(* CODESYS project teltonikaSMSalarmSender.export

Project tree, tasks and I/O mapping:
  libraries: Standard, 3.5.18.0 (System); WagoSysCurl, 1.1.5.0 (WAGO); WagoAppTime, 1.7.3.5 (WAGO); VisuDialogs, * (System)
  task MainTask (cyclic, interval 200 ms, priority 15) calls prg_AlarmSMS
  task VISU_TASK (cyclic, interval 100 ms, priority 15) calls VisuElems.Visu_Prg
  Teltonika/
    global variables GVL_TeltonikaCredentials
    function block FbAlarmSlot [ST]
    function block FbTeltonikaSMS [ST]: ExtractJson
    program prg_AlarmSMS [ST]
  visualisation AlarmAlarms
  visualisation AlarmerListe
  visualisation AlarmMain
*)

// Teltonika/GVL_TeltonikaCredentials
(*
	GVL_TeltonikaCredentials                                  Revised 22.08.2026
	==========================================================================
	WHAT THIS LIST IS FOR
	The single place where the Teltonika router login is maintained. Both the
	older prg_SendSMS and the newer prg_AlarmSMS read from here, so a
	changed password only has to be entered once.

	WHY THE CREDENTIALS ARE RETAIN AND THE REST IS NOT
	Teltonika_Username and Teltonika_Password are VAR_GLOBAL RETAIN, so they
	keep their value through a PLC restart and can be corrected online without
	rebuilding and downloading. That matters because a password change on the
	router would otherwise take a full engineering session to follow.
	The remaining entries are ordinary globals: they belong to the project and
	should come back from the source on every download.

	WHY THE PASSWORD IS BLANK IN THE SOURCE
	So the secret is not stored in the project file, which gets copied, backed
	up and shared. Enter it ONCE online and the retain keeps it.
	If you do decide to put it in the source anyway, remember that the dollar
	sign is the escape character in ST and must be doubled. Ordinary characters
	such as the at sign need no escaping.

	VERIFIED 22.08.2026 ON rutx09-hyc
	The whole API flow - login, modem status returning id 3-1, and send - works
	with the ADMIN user. A separate low privilege user named pfc300 was refused
	with HTTP 401 code 120: it either does not exist on that router, or its user
	group has no API access. To move to a dedicated API user later, create it on
	the correct router, put it in a group allowed to reach the messages
	endpoints, and change the two retain values online. No code change needed.

	Do not publish or share this file.
*)
{attribute 'qualified_only'}
VAR_GLOBAL
	// prg_AlarmSMS therefore overrides the host locally in its own
	// sRouterOverride, and only borrows the credentials from here.
	// Written WITHOUT the https prefix - the send block adds that itself.
	Teltonika_sRouterIP	: STRING := 'rutx09.tailescale.ts.net';

	// Default recipient and message for the older prg_SendSMS. The alarm
	// system does not use these; it keeps its own recipient list.
	Teltonika_Number	: STRING[64] := '+4791919191';
	Teltonika_sMessage	: STRING := 'Debug test SMSCodesys';
END_VAR

VAR_GLOBAL RETAIN
	// Router API user. Must have API rights - an ordinary low privilege user
	// is refused with 401 code 120 even when the password is correct.
	Teltonika_Username	: STRING[64] := 'admin';

	// Blank on purpose, see the note in the header. Enter it online once.
	Teltonika_Password	: STRING[64] := '';
END_VAR

// Teltonika/prg_AlarmSMS
(*
	prg_AlarmSMS                        Created 20.08.2026, rev 23.08.2026
	==========================================================================
	WHAT THIS PROGRAM DOES
	It turns boolean alarm conditions into text messages, and hands them one at
	a time to FbTeltonikaSMS, which talks to a Teltonika RUTX09 router
	over its REST API. The router holds the SIM card, so the PLC needs no modem.

	THE CHAIN, IN ORDER
	  aAlarm[i].xAlarmIn        a condition in the plant becomes TRUE
	  aAlarm[i]                 the slot debounces it and produces xActive plus
	                            the one shot edges xRising and xFalling
	  aAlarm[i].xSmsEnable      the operator switch: may this alarm send at all?
	  aAlarm[i].axToRecipient[] one BOOL per person, picking who gets this alarm
	  aQueueMsg / aQueueNo      a FIFO, because sending takes seconds and alarms
	                            can arrive in bursts
	  oSms                      the router client, driven one message at a time

	WHY EACH ALARM IS A FUNCTION BLOCK INSTANCE
	The CODESYS Best Practices for visualization recommend passing ONE parameter
	to a reusable visualization through VAR_IN_OUT. A slot instance is exactly
	that: a frame showing one row references prg_AlarmSMS.aAlarm[i] and
	gets every field of that alarm with it.

	WHY THE RECIPIENT SELECTION IS AN ARRAY OF BOOL
	Changed 23.08.2026 from a BYTE bit mask. A mask is compact but hostile to a
	visualization: a checkbox has to bind to a single bit, the operator sees a
	meaningless number, and an off by one in the bit index is invisible until
	the wrong person is woken up. One BOOL per recipient binds directly to a
	checkbox and reads the same way in the code.

	WHY A QUEUE AND A RATE LIMIT
	One message needs several task cycles and up to three network round trips.
	Without a queue a burst of alarms would overwrite each other. Without
	iMaxSmsPerHour a chattering signal could send hundreds of messages, which
	costs real money and buries the operator in noise.

	NOTE ON LANGUAGE
	Comments are English. Operator facing texts are deliberately Norwegian,
	because sText goes straight into an SMS that a Norwegian recipient reads.
*)
PROGRAM prg_AlarmSMS
VAR CONSTANT
	// Sizes are constants so the arrays, the loops and the visualization all
	// agree on one number. MAX_RECIPIENTS must match the array size declared
	// inside FbAlarmSlot - raise both together if more than four
	// people need alarms.
	MAX_ALARMS		: INT := 20;	// Alarm slots available for configuration
	MAX_RECIPIENTS	: INT := 4;		// Phone numbers that can receive alarms
	QUEUE_SIZE		: INT := 16;	// Messages that can wait before one is lost
	MAX_RETRY		: INT := 2;		// Extra attempts, and only for KNOWN failures.
									// See the retry policy in section 6 below.
	MSG_MAX_LEN		: INT := 140;	// Message cap. CONCAT returns STRING(255) in
									// CODESYS and the whole JSON body must fit in
									// that, so the text itself is capped here.
END_VAR

VAR
	// =================================================================
	// 1) THE ALARM TABLE
	// -----------------------------------------------------------------
	// One FbAlarmSlot per alarm. Each slot carries its own
	// configuration AND its own live state, and does its own debouncing.
	//
	// Wire your plant conditions into the slots from anywhere in the project:
	//   prg_AlarmSMS.aAlarm[1].xAlarmIn := NOT HTTP_HvaKosterStrommen.xPriceDataValid;
	//
	// A visualization row binds to one whole slot as a single reference:
	//   alarm  ->  prg_AlarmSMS.aAlarm[1]
	//
	// iDelaySec is in SECONDS: 30 is thirty seconds, 120 is two minutes,
	// 300 is five minutes. The slot renders it back as readable text.
	//
	// The recipient selection is NOT set here. Every slot falls back to the
	// default declared in the function block, which is recipient 1 only.
	// Change it per alarm from the visualization, or add axToRecipient to the
	// lines below if a different default suits the plant better.
	//
	// Only slots 1 to 3 are enabled. The rest are written but switched off,
	// because an alarm whose xAlarmIn is not wired yet should not be able to
	// send anything. Enable each one as you connect its signal.
	// =================================================================
	aAlarm : ARRAY[1..MAX_ALARMS] OF FbAlarmSlot := [
		// --- Energi og pris ---
		(xSmsEnable := TRUE,  iDelaySec := 300,
		 sText := 'Stroempriser ikke oppdatert fra hvakosterstrommen.no'),
		(xSmsEnable := TRUE,  iDelaySec := 120,
		 sText := 'Solcelleanlegg: ingen Modbus-kontakt'),
		(xSmsEnable := TRUE,  iDelaySec := 120,
		 sText := 'MQTT-forbindelse mot skyen er nede'),
		(xSmsEnable := FALSE, iDelaySec := 30,
		 sText := 'Hoey stroempris - forbruk boer reduseres'),

		// --- Energimaalere, stigere ---
		(xSmsEnable := FALSE, iDelaySec := 120,
		 sText := 'Energimaaler stiger 433.101 og 433.201 svarer ikke'),
		(xSmsEnable := FALSE, iDelaySec := 120,
		 sText := 'Energimaaler stiger 433.102 og 433.202 svarer ikke'),
		(xSmsEnable := FALSE, iDelaySec := 120,
		 sText := 'Energimaaler stiger 433.103 svarer ikke'),
		(xSmsEnable := FALSE, iDelaySec := 120,
		 sText := 'Energimaaler stiger 433.104 svarer ikke'),
		(xSmsEnable := FALSE, iDelaySec := 120,
		 sText := 'Energimaaler stiger 433.203 svarer ikke'),
		(xSmsEnable := FALSE, iDelaySec := 120,
		 sText := 'Energimaaler stiger 434.001 svarer ikke'),

		// --- Varme ---
		(xSmsEnable := FALSE, iDelaySec := 120,
		 sText := 'Elkjele: ingen kontakt med energimaaler'),
		(xSmsEnable := FALSE, iDelaySec := 120,
		 sText := 'Varmepumpe: ingen kontakt med energimaaler'),

		// --- Ventilasjon ---
		(xSmsEnable := FALSE, iDelaySec := 120,
		 sText := 'Ventilasjonsaggregat 360.003 svarer ikke'),
		(xSmsEnable := FALSE, iDelaySec := 120,
		 sText := 'Ventilasjonsaggregat 360.004 svarer ikke'),
		(xSmsEnable := FALSE, iDelaySec := 120,
		 sText := 'Ventilasjonsaggregat 360.005 svarer ikke'),

		// --- Varmtvann og feltbuss ---
		(xSmsEnable := FALSE, iDelaySec := 120,
		 sText := 'Varmtvannsbereder CH124 svarer ikke'),
		(xSmsEnable := FALSE, iDelaySec := 60,
		 sText := 'Modbus RTU-linje 1: kommunikasjonsfeil'),
		(xSmsEnable := FALSE, iDelaySec := 120,
		 sText := 'Teltonika-ruter: ingen Modbus-kontakt'),

		// --- Reserve ---
		(xSmsEnable := FALSE, iDelaySec := 30,
		 sText := 'Reserve - ledig alarmplass 19'),
		(xSmsEnable := FALSE, iDelaySec := 30,
		 sText := 'Reserve - ledig alarmplass 20')];

	// =================================================================
	// 2) RECIPIENTS
	// -----------------------------------------------------------------
	// Three parallel arrays, index 1 to 4. A recipient must be enabled here
	// AND selected in the slot before anything is sent, so one person can be
	// taken out of service without editing every alarm.
	//
	// In a visualization, bind a CHECKBOX to axRecipientEnable[n], and text
	// fields with %s to the name and the number.
	// =================================================================
	axRecipientEnable	: ARRAY[1..MAX_RECIPIENTS] OF BOOL       := [TRUE, FALSE, FALSE, FALSE];	// On or off per person
	asRecipientName		: ARRAY[1..MAX_RECIPIENTS] OF STRING(20) := ['Espen', '', '', ''];			// Display only, never sent
	asRecipientNumber	: ARRAY[1..MAX_RECIPIENTS] OF STRING(24) := ['+4791916159', '', '', ''];	// International format, this is what is dialled

	// =================================================================
	// 3) GENERAL SETTINGS
	// =================================================================
	xSmsGlobalEnable	: BOOL := TRUE;			// Master switch. FALSE stops all sending and all
												// queueing - use it during service work.
	xSendOkMessages		: BOOL := TRUE;			// Also send a message when an alarm clears, so the
												// operator knows the fault went away.
	sSiteName			: STRING(20) := 'PFC300';	// Prefix in every message. Essential when one
												// phone receives alarms from several plants.
	iMaxSmsPerHour		: INT := 15;			// Hard ceiling per rolling hour, against runaway cost
	tPauseBetweenSms	: TIME := T#10S;		// Gap between messages. Gives the router time to hand
												// the previous one over, and guarantees a clean edge.
	tRetryDelay			: TIME := T#60S;		// Wait before repeating a message that failed for a
												// known reason, so a brief outage can recover.

	// Leave EMPTY to fall back
	// to GVL_TeltonikaCredentials.Teltonika_sRouterIP.
	sRouterOverride		: STRING(80) := '';

	// Modem id inside the router. Leave EMPTY for auto-detection, which is
	// normal and survives the id changing after a router restart.
	sModemIdForced		: STRING(16) := '';

	// =================================================================
	// STATUS AND DIAGNOSTICS
	// -----------------------------------------------------------------
	// Read only. These exist to be bound to a visualization, and to make a
	// failure explain itself without a debugger attached.
	// =================================================================
	sRouterInUse			: STRING(80);	// Host actually used, after the override is resolved
	xCredentialsMissing		: BOOL;			// TRUE when user name or password is blank. Blocks
											// sending so the queue is not burned on doomed logins.
	iQueueCount				: INT;			// Messages waiting right now
	xRateLimited			: BOOL;			// TRUE when the hourly ceiling holds messages back
	iSentThisHour			: INT;			// Counter behind the ceiling, reset once an hour
	iEnabledCount			: INT;			// How many of the twenty alarms are switched on. Handy
											// as a single number on an overview screen.
	iActiveCount			: INT;			// How many alarms are standing right now
	udiSentOk				: UDINT;		// Messages the router confirmed, since PLC start
	udiSendFailed			: UDINT;		// Messages given up on after all allowed retries
	udiUncertain			: UDINT;		// Messages whose fate is unknown - the request went out
											// but no answer came back. Never retried, to avoid
											// sending the same SMS twice.
	udiDropped				: UDINT;		// Messages never queued because the FIFO was full
	sLastMessage			: STRING(140);	// Exact text last handed to the router
	sLastError				: STRING(200);	// Why the last attempt failed
	sSmsStatus				: STRING(200);	// Live progress text from the send FB
	sCurlError				: STRING(200);	// Raw libcurl error. The one to read when diHttpCode
											// stays 0, because then there is no HTTP answer.
	diHttpCode				: DINT;			// HTTP status of the last request. 0 means the request
											// never produced an HTTP answer at all.
	uiSendStep				: UINT;			// Live step inside the send FB: 10 and 11 login,
											// 20 and 21 modem lookup, 30 and 31 the send itself.

	// =================================================================
	// MANUAL TEST
	// -----------------------------------------------------------------
	// One button, two destinations. Leave sTestNumber EMPTY and the test goes
	// to every enabled recipient, which proves the real alarm path end to end.
	// Type a number into sTestNumber and it goes only there, which is how you
	// check a new phone before adding it to the recipient list.
	// xManualSend is self resetting, so a visualization button only has to
	// toggle it and the program clears it again on the next cycle.
	// =================================================================
	xManualSend			: BOOL;								// Set TRUE to queue one test message
	sTestNumber			: STRING(24) := '';					// Optional. Empty means all enabled recipients.
	sManualText			: STRING(100) := 'Testmelding fra PFC300';	// Body of the test message
	iTestQueued			: INT;								// How many messages the last test queued,
															// so the operator sees it did something

	// =================================================================
	// INTERNALS - not intended for the visualization
	// =================================================================
	aQueueMsg			: ARRAY[1..QUEUE_SIZE] OF STRING(140);	// FIFO slot: the message text
	aQueueNo			: ARRAY[1..QUEUE_SIZE] OF STRING(24);	// FIFO slot: the recipient number.
																// Kept beside the text so one alarm
																// to three people becomes three
																// independent queue entries.
	iQHead				: INT;					// Last slot read from, wraps at QUEUE_SIZE
	iQTail				: INT;					// Last slot written to, wraps at QUEUE_SIZE

	oSms				: FbTeltonikaSMS;	// The router client. Called every cycle so its
													// asynchronous transfer can advance.
	xSendTrigger		: BOOL;					// Rising edge starts oSms. Held TRUE for the whole
												// job and cleared afterwards, so the next message
												// gets a fresh edge.
	iSendState			: INT;					// Sender state machine, see section 6
	iRetry				: INT;					// Attempts already used on the current message
	sCurMsg				: STRING(140);			// The message being sent right now
	sCurNo				: STRING(24);			// The recipient it is going to

	TON_Pause			: TON;					// Enforces tPauseBetweenSms between messages
	TON_Retry			: TON;					// Enforces tRetryDelay before a repeat attempt
	TON_HourWindow		: TON;					// Free running one hour timer that clears
												// iSentThisHour, implementing the rate limit

	xManualPrev			: BOOL;					// Edge memory for xManualSend
	i					: INT;					// Loop counter over the alarm slots
	iRcp				: INT;					// Loop counter over the recipients. NOTE: a bare
												// r cannot be used as an identifier - CODESYS
												// reserves R and S as the IL reset and set
												// operators, and the parser fails cryptically.
	iGuard				: INT;					// Safety counter so the sanitize loop can never
												// spin forever on malformed text
	iQuote				: INT;					// Position of the next double quote to remove
	xQueueIt			: BOOL;					// Set when the slot being scanned needs sending
	sMsg				: STRING(140);			// Message being assembled
	sStamp				: STRING(30);			// Time stamp for the message, format dd.mm hh:mm
	sRaw				: STRING(40);			// Raw DT_TO_STRING output the stamp is cut from
END_VAR

// =====================================================================
// 1) Resolve which router host to talk to.
//    The local override wins, or if it is emty use so GVL_TeltonikaCredentials.Teltonika_sRouterIP
// =====================================================================
IF LEN(sRouterOverride) > 0 THEN
	sRouterInUse := sRouterOverride;
ELSE
	sRouterInUse := GVL_TeltonikaCredentials.Teltonika_sRouterIP;
END_IF

// Without credentials every login is doomed, and each doomed attempt costs a
// network round trip and fills the diagnostics with noise. Detect it once here
// and let section 6 hold the queue instead.
xCredentialsMissing := (LEN(GVL_TeltonikaCredentials.Teltonika_Username) = 0)
					OR (LEN(GVL_TeltonikaCredentials.Teltonika_Password) = 0);

// =====================================================================
// 2) Rolling one hour window behind the rate limit.
//    A free running timer is enough: it does not matter exactly where the
//    hour boundary falls, only that the counter cannot grow forever.
// =====================================================================
TON_HourWindow(IN := TRUE, PT := T#1H);
IF TON_HourWindow.Q THEN
	TON_HourWindow(IN := FALSE);	// Restart the window
	iSentThisHour := 0;
END_IF

// =====================================================================
// 3) Build the time stamp that goes into every message.
//    DT_TO_STRING has a fixed layout, so the parts can be cut out by
//    position instead of parsed:
//        DT#2026-08-20-14:20:28
//            ^4      ^9 ^12 ^15
// =====================================================================
sRaw   := DT_TO_STRING(WagoAppTime.FuGetLocalDateAndTime());
sStamp := CONCAT(MID(sRaw, 2, 12), '.');		// Two digits of day
sStamp := CONCAT(sStamp, MID(sRaw, 2, 9));		// Two digits of month
sStamp := CONCAT(sStamp, ' ');
sStamp := CONCAT(sStamp, MID(sRaw, 5, 15));		// Five characters, hh:mm

// =====================================================================
// 4) Scan every alarm slot and queue messages for the transitions.
//    Calling the slot updates its debounce timer and its edge outputs, so
//    all the per alarm timing logic lives in the slot rather than here.
//    Only transitions produce messages: a standing alarm stays silent.
// =====================================================================
iEnabledCount := 0;
iActiveCount  := 0;

FOR i := 1 TO MAX_ALARMS DO

	aAlarm[i]();			// Debounce and edge detection happen inside the slot
	xQueueIt := FALSE;

	// Two counters for the overview screen, so the operator can see at a
	// glance how much of the system is armed and how much is in alarm.
	IF aAlarm[i].xSmsEnable THEN
		iEnabledCount := iEnabledCount + 1;
	END_IF
	IF aAlarm[i].xActive THEN
		iActiveCount := iActiveCount + 1;
	END_IF

	IF xSmsGlobalEnable AND aAlarm[i].xSmsEnable THEN
		IF aAlarm[i].xRising THEN
			// The alarm has just appeared.
			sMsg     := CONCAT(sSiteName, ' ');
			sMsg     := CONCAT(sMsg, sStamp);
			sMsg     := CONCAT(sMsg, ' ALARM: ');
			sMsg     := CONCAT(sMsg, aAlarm[i].sText);
			xQueueIt := TRUE;
		ELSIF aAlarm[i].xFalling AND xSendOkMessages THEN
			// The alarm has cleared. Optional, because on a noisy signal this
			// doubles the number of messages.
			sMsg     := CONCAT(sSiteName, ' ');
			sMsg     := CONCAT(sMsg, sStamp);
			sMsg     := CONCAT(sMsg, ' OK: ');
			sMsg     := CONCAT(sMsg, aAlarm[i].sText);
			xQueueIt := TRUE;
		END_IF
	END_IF

	IF xQueueIt THEN
		// The message is embedded in a JSON body, where a double quote would
		// end the string early and corrupt the request. Replace any with
		// spaces. The guard counter bounds the loop so malformed text can
		// never stall the task.
		iGuard := 0;
		iQuote := FIND(sMsg, '"');
		WHILE (iQuote > 0) AND (iGuard < 20) DO
			sMsg   := REPLACE(sMsg, ' ', 1, iQuote);
			iQuote := FIND(sMsg, '"');
			iGuard := iGuard + 1;
		END_WHILE

		IF LEN(sMsg) > MSG_MAX_LEN THEN
			sMsg := LEFT(sMsg, MSG_MAX_LEN);
		END_IF

		// One queue entry per selected recipient. Two conditions have to agree:
		// the person must be in service at all (axRecipientEnable) AND this
		// particular alarm must be addressed to them (axToRecipient). Queueing
		// per recipient rather than per alarm keeps the sender simple: it never
		// has to know that one alarm can have several destinations.
		FOR iRcp := 1 TO MAX_RECIPIENTS DO
			IF axRecipientEnable[iRcp]
				AND aAlarm[i].axToRecipient[iRcp]
				AND (LEN(asRecipientNumber[iRcp]) > 0) THEN

				IF iQueueCount < QUEUE_SIZE THEN
					iQTail            := (iQTail MOD QUEUE_SIZE) + 1;	// Ring buffer wrap
					aQueueMsg[iQTail] := sMsg;
					aQueueNo[iQTail]  := asRecipientNumber[iRcp];
					iQueueCount       := iQueueCount + 1;
				ELSE
					// Queue full. Counting the loss is better than blocking the
					// task or discarding it unnoticed.
					udiDropped := udiDropped + 1;
				END_IF
			END_IF
		END_FOR
	END_IF
END_FOR

// =====================================================================
// 5) Manual test message.
//    Two destinations from one button:
//      sTestNumber empty     -> every enabled recipient, which proves the
//                               real alarm path exactly as an alarm would use it
//      sTestNumber filled in -> only that number, for checking a new phone
//                               before it is added to the recipient list
//    iTestQueued reports back how many messages were actually queued, so a
//    press that produced nothing is visible rather than silent.
// =====================================================================
IF xManualSend AND NOT xManualPrev THEN
	sMsg := CONCAT(sSiteName, ' ');
	sMsg := CONCAT(sMsg, sStamp);
	sMsg := CONCAT(sMsg, ' TEST: ');
	sMsg := CONCAT(sMsg, sManualText);

	// Same sanitizing as a real alarm, because the operator types this text
	// and a double quote would corrupt the JSON body just the same.
	iGuard := 0;
	iQuote := FIND(sMsg, '"');
	WHILE (iQuote > 0) AND (iGuard < 20) DO
		sMsg   := REPLACE(sMsg, ' ', 1, iQuote);
		iQuote := FIND(sMsg, '"');
		iGuard := iGuard + 1;
	END_WHILE

	IF LEN(sMsg) > MSG_MAX_LEN THEN
		sMsg := LEFT(sMsg, MSG_MAX_LEN);
	END_IF

	iTestQueued := 0;

	IF LEN(sTestNumber) > 0 THEN
		// A number was typed in, so send only there.
		IF iQueueCount < QUEUE_SIZE THEN
			iQTail            := (iQTail MOD QUEUE_SIZE) + 1;
			aQueueMsg[iQTail] := sMsg;
			aQueueNo[iQTail]  := sTestNumber;
			iQueueCount       := iQueueCount + 1;
			iTestQueued       := 1;
		ELSE
			udiDropped := udiDropped + 1;
		END_IF
	ELSE
		// No number typed, so send to everyone who is enabled - the same set
		// an alarm addressed to all four recipients would reach.
		FOR iRcp := 1 TO MAX_RECIPIENTS DO
			IF axRecipientEnable[iRcp] AND (LEN(asRecipientNumber[iRcp]) > 0) THEN
				IF iQueueCount < QUEUE_SIZE THEN
					iQTail            := (iQTail MOD QUEUE_SIZE) + 1;
					aQueueMsg[iQTail] := sMsg;
					aQueueNo[iQTail]  := asRecipientNumber[iRcp];
					iQueueCount       := iQueueCount + 1;
					iTestQueued       := iTestQueued + 1;
				ELSE
					udiDropped := udiDropped + 1;
				END_IF
			END_IF
		END_FOR
	END_IF
END_IF
xManualPrev := xManualSend;
xManualSend := FALSE;			// Clear it again so the button is momentary

// =====================================================================
// 6) The sender.
//    Strictly one message at a time. The send FB can only handle one job, and
//    serialising here also means the router is never hit by parallel requests.
//
//    RETRY POLICY, and why it is not simply MAX_RETRY attempts:
//    Repeating a request is only safe when we KNOW nothing was sent. A login
//    failure, or a rejection carrying a real HTTP status, both mean the router
//    did nothing, so those are retried. But if the send request went out and
//    no answer came back, the router may already have queued the SMS -
//    repeating it would deliver the same message twice. The send FB flags that
//    case with xSendUncertain, and such a message is dropped and counted.
// =====================================================================
CASE iSendState OF

	// -----------------------------------------------------------------
	0:	// Idle. Take the next message out of the queue if everything allows it.
	// -----------------------------------------------------------------
		xSendTrigger := FALSE;
		xRateLimited := (iSentThisHour >= iMaxSmsPerHour) AND (iQueueCount > 0);

		IF (iQueueCount > 0)
			AND xSmsGlobalEnable
			AND NOT xRateLimited
			AND NOT xCredentialsMissing THEN

			iQHead      := (iQHead MOD QUEUE_SIZE) + 1;		// Ring buffer wrap
			sCurMsg     := aQueueMsg[iQHead];
			sCurNo      := aQueueNo[iQHead];
			iQueueCount := iQueueCount - 1;
			iRetry      := 0;
			iSendState  := 10;
		END_IF

	// -----------------------------------------------------------------
	10:	// Start one attempt. Raising xSendTrigger gives the send FB the rising
	//     edge it needs; it stays TRUE until the job finishes.
	// -----------------------------------------------------------------
		sLastMessage := sCurMsg;
		xSendTrigger := TRUE;
		iSendState   := 20;

	// -----------------------------------------------------------------
	20:	// Wait for the verdict. The send FB is asynchronous and advances one
	//     step per call, so this state is held for several cycles.
	// -----------------------------------------------------------------
		IF oSms.xDone THEN
			xSendTrigger  := FALSE;
			udiSentOk     := udiSentOk + 1;
			iSentThisHour := iSentThisHour + 1;
			iSendState    := 30;

		ELSIF oSms.xError THEN
			xSendTrigger := FALSE;
			sLastError   := oSms.sErrorText;

			IF oSms.xSendUncertain THEN
				// Unknown outcome, see the retry policy above. The hour slot is
				// counted as used as well, because the message probably did cost
				// an SMS and the rate limit should not underestimate usage.
				udiUncertain  := udiUncertain + 1;
				iSentThisHour := iSentThisHour + 1;
				iSendState    := 30;

			ELSIF iRetry < MAX_RETRY THEN
				// Known failure, nothing was sent, so trying again is safe.
				iRetry     := iRetry + 1;
				iSendState := 40;

			ELSE
				// Out of attempts. Give up on this one and move on, rather than
				// letting a single bad message block the whole queue.
				udiSendFailed := udiSendFailed + 1;
				iSendState    := 30;
			END_IF
		END_IF

	// -----------------------------------------------------------------
	30:	// Pause between messages. Two purposes: breathing room for the router,
	//     and it guarantees at least one cycle with xSendTrigger FALSE so the
	//     next message produces a genuine rising edge.
	// -----------------------------------------------------------------
		TON_Pause(IN := TRUE, PT := tPauseBetweenSms);
		IF TON_Pause.Q THEN
			TON_Pause(IN := FALSE);
			iSendState := 0;
		END_IF

	// -----------------------------------------------------------------
	40:	// Wait before repeating the same message, so a brief outage has time
	//     to clear instead of burning all attempts in a few seconds.
	// -----------------------------------------------------------------
		TON_Retry(IN := TRUE, PT := tRetryDelay);
		IF TON_Retry.Q THEN
			TON_Retry(IN := FALSE);
			iSendState := 10;
		END_IF

ELSE
	// Unknown state. Reached only after an online change moves the code under
	// a running state machine. Returning to idle is always safe.
	iSendState := 0;
END_CASE

// =====================================================================
// 7) Call the router client.
//    This MUST run every cycle, including when idle: the underlying cURL
//    transfer is asynchronous and only advances when the FB body executes.
// =====================================================================
oSms(
	sRouterIP      := sRouterInUse,
	sUsername      := GVL_TeltonikaCredentials.Teltonika_Username,
	sPassword      := GVL_TeltonikaCredentials.Teltonika_Password,
	sNumber        := sCurNo,
	sMessage       := sCurMsg,
	sModemIdForced := sModemIdForced,
	xSend          := xSendTrigger);

// Mirror the interesting outputs so a visualization can bind them here rather
// than reaching into the FB instance. Everything else is still reachable as
// oSms.<name>, for example oSms.udiLoginCnt and oSms.xTokenValid.
sSmsStatus := oSms.sStatus;
sCurlError := oSms.sCurlError;		// The one that explains a diHttpCode of 0
diHttpCode := oSms.diHttpCode;
uiSendStep := oSms.uiStepOut;		// 10 and 11 login, 20 and 21 modem, 30 and 31 send

END_PROGRAM

// Teltonika/FbTeltonikaSMS
(*
	FbTeltonikaSMS                      Created 20.08.2026, rev 22.08.2026
	==========================================================================
	WHAT THIS BLOCK DOES
	Sends ONE text message through a Teltonika RUTX router using its REST API.
	The router holds the SIM card, so the PLC needs no modem. Give it a number
	and a text, pulse xSend, and watch xDone or xError.

	Reference implementation: github.com/espenbo/wagoEdgeStart/TeltonikaRouter
	and the working /root/sendsms_busyboxV3.sh on this PLC. Both were used to
	prove the API flow before it was written in ST.

	THE API FLOW - THREE REQUESTS
	  1  POST /api/login                 user and password  ->  bearer token
	  2  GET  /api/modems/status         token              ->  modem id, 3-1 here
	  3  POST /api/messages/actions/send token, number, text, modem id
	The router answers the third with success true when it has accepted the SMS.

	*** WHY EVERY REQUEST IS SPLIT IN TWO STEPS ***
	WagoSysCurl.FbCurl is ASYNCHRONOUS. curl_easy_perform() only STARTS the
	transfer and returns immediately; the FB reports progress through xBusy,
	xDone and xError, and its body must be called every cycle for those to
	update. Reading curl_easy_getResponseCode() straight after perform therefore
	always yields 0 and an empty receive buffer - which looks exactly like a
	network failure and is extremely misleading. Each request is consequently a
	start step followed by a wait step:

	  10 login start   11 login wait
	  20 modem start   21 modem wait
	  30 send start    31 send wait
	 100 done         900 error

	Every wait step is bounded by tWaitTimeout, so a transfer that never
	completes cannot freeze the state machine.

	*** TOKEN CACHING ***
	The router reports expires 299, so a token is good for just under five
	minutes. Both the token and the detected modem id survive between messages,
	so a follow up message jumps straight to step 30: two steps and one network
	round trip instead of eight steps and three. If the router rejects a cached
	token with HTTP 401 the block logs in again once and repeats the request,
	which is safe because a 401 proves nothing was sent.

	*** DUPLICATE PROTECTION ***
	If the send request goes out and no answer comes back, the router may
	already have accepted the SMS. Repeating it would deliver the same message
	twice. That case raises xSendUncertain, and the caller must not retry while
	it is set. A clean HTTP answer reporting failure is safe to repeat.

	*** LENGTH LIMITS TO RESPECT ***
	CONCAT returns STRING(255) in CODESYS, so the assembled JSON body cannot
	exceed that. sMessage is therefore capped at 140 characters, which also
	keeps the SMS inside a single 160 character GSM message.
*)
FUNCTION_BLOCK FbTeltonikaSMS
VAR_INPUT
	// --- What to send, and where ---
	sRouterIP		: STRING(80);		// Router host name or IP. WITHOUT the https prefix,
										// the block adds that when building the URL.
	sUsername		: STRING(64);		// Router API user. Must have API rights - an ordinary
										// low privilege user is rejected with 401 code 120.
	sPassword		: STRING(64);		// Password for that user
	sNumber			: STRING(32);		// Recipient, international format, for example +47...
	sMessage		: STRING(140);		// The text itself. See the length note in the header.

	// --- Behaviour tuning ---
	sModemIdForced	: STRING(16) := '';	// Leave EMPTY for auto-detection, which is normal and
										// survives the id changing after a router restart.
										// Set it only to pin one specific modem.
	tRequestTimeout	: TIME := T#15S;	// Passed down to cURL as its own transfer timeout
	tWaitTimeout	: TIME := T#30S;	// Guard in the wait steps. Keep it LONGER than
										// tRequestTimeout, so cURL gets to fail on its own
										// terms first and can report a proper reason.
	tTokenLifetime	: TIME := T#4M;		// How long a token is reused before logging in again.
										// The router says 299 s, so stay safely below that.

	// --- Control ---
	xSend			: BOOL;				// RISING EDGE starts one send job. Level is ignored
										// while a job is already running.
END_VAR
VAR_OUTPUT
	// --- Job state ---
	xBusy			: BOOL;				// TRUE from the rising edge until done or failed
	xDone			: BOOL;				// Latched TRUE when the router confirmed the SMS.
										// Cleared when the next job starts.
	xError			: BOOL;				// Latched TRUE when the job failed. Read sErrorText.
	xSendUncertain	: BOOL;				// TRUE when the SMS may or may not have gone out.
										// The caller MUST NOT retry the message while set,
										// or the recipient can receive it twice.
	xTokenValid		: BOOL;				// TRUE while a cached token can still be reused

	// --- Human readable status ---
	sErrorText		: STRING(200);		// Why the last job failed, including HTTP code and,
										// where useful, the raw answer from the router
	sStatus			: STRING(200);		// Live progress text, useful on a visualization
	tLastSend		: DT;				// Time stamp of the last confirmed send

	// --- Counters, all since PLC start ---
	sModemID		: STRING(16);		// Modem id currently in use. Kept between messages so
										// the lookup runs once rather than every time.
	udiSentCnt		: UDINT;			// Messages the router confirmed
	udiErrorCnt		: UDINT;			// Jobs that ended in failure
	udiLoginCnt		: UDINT;			// Actual logins performed. Compare with udiSentCnt to
										// see token caching working: it should stay well below.

	// --- Raw diagnostics from the last completed request ---
	diHttpCode		: DINT;				// HTTP status. 0 is special: it means the transfer
										// never produced an HTTP answer at all, so look at
										// sCurlError instead of trying to interpret the code.
	xCurlError		: BOOL;				// libcurl reported a transport level error
	sCurlError		: STRING(200);		// libcurl error text. The real explanation whenever
										// diHttpCode is 0, for example a name resolution
										// failure or an SSL connect error.
	sCurlSource		: STRING(100);		// Where inside libcurl the error came from
	sLastResponse	: STRING(200);		// First 200 characters of the router answer, so a
										// rejection can be read without a network trace
	uiStepOut		: UINT;				// Mirror of the internal step, for commissioning
END_VAR
VAR
	fbCurl			: WagoSysCurl.FbCurl;	// The cURL handle. ASYNCHRONOUS - see header.
	uiStep			: UINT;				// State machine position, see the header for the map
	xSendPrev		: BOOL;				// Edge memory for xSend
	TON_Wait		: TON;				// Bounds each wait step, so a stalled transfer cannot
										// hold the state machine forever
	TON_TokenAge	: TON;				// Ages the cached token out after tTokenLifetime
	xRetriedLogin	: BOOL;				// Allows exactly ONE forced re-login per job after a
										// 401, so a stale token cannot cause an endless loop
	sResponse		: STRING(4095);		// Receive buffer for the HTTP body. Deliberately large:
										// the modem status answer carries many fields.
	sURL			: STRING(200);		// Assembled request URL
	sBody			: STRING(254);		// Assembled JSON request body. Sized just under the
										// 255 characters CONCAT can produce.
	sHeader			: STRING(250);		// Assembled Authorization header
	sToken			: STRING(200);		// Bearer token. Reused across messages until it ages
										// out or the router rejects it.
END_VAR

// =====================================================================
// The FB body must run EVERY cycle, idle or not. The cURL transfer is
// asynchronous and only makes progress when this executes; skipping it
// would leave xBusy, xDone and xError frozen at their old values.
// =====================================================================
fbCurl();
uiStepOut := uiStep;

// =====================================================================
// Age the cached token out.
// The timer runs only while a token is held, so it measures the age of that
// specific token. When it expires the token is discarded and the next job
// logs in again. tTokenLifetime sits below the 299 seconds the router
// reports, so we never present a token the router has already forgotten.
// =====================================================================
TON_TokenAge(IN := xTokenValid, PT := tTokenLifetime);
IF TON_TokenAge.Q THEN
	xTokenValid := FALSE;
	sToken      := '';
END_IF

// =====================================================================
// A rising edge on xSend starts one job. A job in progress is never
// interrupted, so a caller cannot corrupt a transfer by pulsing again.
//
// The entry point depends on what is still cached. With a valid token and a
// known modem id the job starts directly at the send step, which is the whole
// point of the caching: two steps instead of eight.
// =====================================================================
IF xSend AND NOT xSendPrev AND NOT xBusy THEN
	xBusy          := TRUE;
	xDone          := FALSE;
	xError         := FALSE;
	xSendUncertain := FALSE;
	xRetriedLogin  := FALSE;	// Fresh job, so the one allowed re-login is available again
	sErrorText     := '';
	diHttpCode     := 0;

	IF xTokenValid AND (LEN(sToken) > 0) THEN
		IF LEN(sModemIdForced) > 0 THEN
			sModemID := sModemIdForced;
			uiStep   := 30;		// Token cached and modem pinned by the operator
		ELSIF LEN(sModemID) > 0 THEN
			uiStep   := 30;		// Token cached and modem detected earlier
		ELSE
			uiStep   := 20;		// Token cached but the modem is still unknown
		END_IF
	ELSE
		uiStep := 10;			// No usable token, so start with a login
	END_IF
END_IF
xSendPrev := xSend;

// =====================================================================
// The state machine.
//
// libcurl option numbers used below, since the WAGO wrapper takes raw ints:
//   13 = TIMEOUT in seconds     47 = POST             64 = SSL_VERIFYPEER
//   78 = CONNECTTIMEOUT         80 = HTTPGET          81 = SSL_VERIFYHOST
//   10002 = URL   10015 = POSTFIELDS   10018 = USERAGENT   10023 = HTTPHEADER
//
// Certificate checking is switched off because the router presents a self
// signed certificate that no public CA vouches for. That is acceptable here
// because the traffic already runs inside the Tailscale tunnel, which does
// its own authentication and encryption.
// =====================================================================
CASE uiStep OF

	// -----------------------------------------------------------------
	0:	// Idle, waiting for a rising edge on xSend.
	// -----------------------------------------------------------------
		xBusy := FALSE;

	// -----------------------------------------------------------------
	10:	// LOGIN - start the request.
	//     Any previous token is dropped first, so a failure here cannot leave
	//     a half valid credential behind for the next job to trip over.
	// -----------------------------------------------------------------
		sStatus     := 'Steg 10: logger inn paa ruteren...';
		sResponse   := '';
		xTokenValid := FALSE;
		sToken      := '';

		fbCurl.curl_easy_init();
		fbCurl.curl_set_RAM(ADR(sResponse), SIZEOF(sResponse));		// Where the answer lands
		fbCurl.curl_easy_setopt_BOOL(64, FALSE);					// Do not verify the certificate
		fbCurl.curl_easy_setopt_BOOL(81, FALSE);					// Do not verify the host name
		fbCurl.curl_easy_setopt_DINT(13, TIME_TO_DINT(tRequestTimeout) / 1000);
		fbCurl.curl_easy_setopt_DINT(78, 10);						// Connect timeout, seconds
		fbCurl.curl_easy_setopt_DINT(47, 1);						// This is a POST

		sURL := CONCAT('https://', sRouterIP);
		sURL := CONCAT(sURL, '/api/login');
		fbCurl.curl_easy_setopt_STRING(10002, sURL);

		// The API only accepts JSON, so the content type has to be declared.
		fbCurl.curl_slist_append(1, 'Content-Type: application/json');
		fbCurl.curl_easy_setopt_slist(10023, 1);

		sBody := CONCAT('{"username":"', sUsername);
		sBody := CONCAT(sBody, '","password":"');
		sBody := CONCAT(sBody, sPassword);
		sBody := CONCAT(sBody, '"}');
		fbCurl.curl_easy_setopt_STRING(10015, sBody);

		fbCurl.curl_easy_perform();		// Starts the transfer and returns at once
		TON_Wait(IN := FALSE);			// Arm the guard timer for the wait step
		uiStep := 11;

	// -----------------------------------------------------------------
	11:	// LOGIN - wait for the answer, then pull the token out of it.
	// -----------------------------------------------------------------
		TON_Wait(IN := TRUE, PT := tWaitTimeout);
		IF fbCurl.xDone OR fbCurl.xError THEN
			TON_Wait(IN := FALSE);

			// Capture everything libcurl knows BEFORE cleaning the handle up,
			// otherwise the diagnostics are lost with it.
			diHttpCode    := LINT_TO_DINT(fbCurl.curl_easy_getResponseCode());
			xCurlError    := fbCurl.xError;
			sCurlError    := fbCurl.sErrorString;
			sCurlSource   := fbCurl.sErrorSource;
			sLastResponse := LEFT(sResponse, 200);

			// Free the header list and the handle. Skipping this leaks memory
			// and lets headers accumulate across requests.
			fbCurl.curl_slist_free_all(1);
			fbCurl.curl_easy_cleanup();

			sToken := ExtractJson(sSource := sResponse, sKey := '"token"');
			IF LEN(sToken) > 0 THEN
				xTokenValid := TRUE;			// Also starts the token age timer
				udiLoginCnt := udiLoginCnt + 1;
				sStatus     := 'Token mottatt';
				IF LEN(sModemIdForced) > 0 THEN
					sModemID := sModemIdForced;
					uiStep   := 30;
				ELSIF LEN(sModemID) > 0 THEN
					uiStep   := 30;
				ELSE
					uiStep   := 20;
				END_IF
			ELSE
				// No token in the answer. Report the HTTP code, and add whichever
				// detail actually explains it: the router answer when there is
				// one, the libcurl reason when the transfer never got that far.
				sErrorText := CONCAT('Innlogging feilet, HTTP ', DINT_TO_STRING(diHttpCode));
				IF diHttpCode = 0 THEN
					sErrorText := CONCAT(sErrorText, ' curl: ');
					sErrorText := CONCAT(sErrorText, LEFT(sCurlError, 110));
				ELSE
					sErrorText := CONCAT(sErrorText, ' svar: ');
					sErrorText := CONCAT(sErrorText, LEFT(sResponse, 110));
				END_IF
				uiStep := 900;
			END_IF

		ELSIF TON_Wait.Q THEN
			// The transfer never reported completion. Abort it explicitly so
			// libcurl releases the connection instead of leaving it dangling.
			TON_Wait(IN := FALSE);
			fbCurl.curl_easy_abort();
			fbCurl.curl_slist_free_all(1);
			fbCurl.curl_easy_cleanup();
			sErrorText := 'Tidsavbrudd under innlogging';
			uiStep     := 900;
		END_IF

	// -----------------------------------------------------------------
	20:	// MODEM ID - start the request.
	//     The send endpoint needs to know which modem to use, and the id is
	//     not fixed: it depends on the hardware slot and can change after a
	//     router restart. Asking is more robust than hard coding.
	// -----------------------------------------------------------------
		sStatus   := 'Steg 20: henter modem-ID...';
		sResponse := '';

		fbCurl.curl_easy_init();
		fbCurl.curl_set_RAM(ADR(sResponse), SIZEOF(sResponse));
		fbCurl.curl_easy_setopt_BOOL(64, FALSE);
		fbCurl.curl_easy_setopt_BOOL(81, FALSE);
		fbCurl.curl_easy_setopt_DINT(13, TIME_TO_DINT(tRequestTimeout) / 1000);
		fbCurl.curl_easy_setopt_DINT(78, 10);
		fbCurl.curl_easy_setopt_DINT(80, 1);						// This one is a GET

		sURL := CONCAT('https://', sRouterIP);
		sURL := CONCAT(sURL, '/api/modems/status');
		fbCurl.curl_easy_setopt_STRING(10002, sURL);

		// Everything past the login is authenticated with the bearer token.
		sHeader := CONCAT('Authorization: Bearer ', sToken);
		fbCurl.curl_slist_append(1, sHeader);
		fbCurl.curl_easy_setopt_slist(10023, 1);

		fbCurl.curl_easy_perform();
		TON_Wait(IN := FALSE);
		uiStep := 21;

	// -----------------------------------------------------------------
	21:	// MODEM ID - wait, then take the first id the router reports.
	// -----------------------------------------------------------------
		TON_Wait(IN := TRUE, PT := tWaitTimeout);
		IF fbCurl.xDone OR fbCurl.xError THEN
			TON_Wait(IN := FALSE);

			diHttpCode    := LINT_TO_DINT(fbCurl.curl_easy_getResponseCode());
			xCurlError    := fbCurl.xError;
			sCurlError    := fbCurl.sErrorString;
			sCurlSource   := fbCurl.sErrorSource;
			sLastResponse := LEFT(sResponse, 200);

			fbCurl.curl_slist_free_all(1);
			fbCurl.curl_easy_cleanup();

			IF (diHttpCode = 401) AND NOT xRetriedLogin THEN
				// The cached token was refused, most likely because the router
				// restarted. Nothing was sent, so logging in again and repeating
				// this request is safe. Allowed only once per job.
				xTokenValid   := FALSE;
				sToken        := '';
				xRetriedLogin := TRUE;
				sStatus       := 'Token avvist - logger inn paa nytt';
				uiStep        := 10;
			ELSE
				sModemID := ExtractJson(sSource := sResponse, sKey := '"id"');
				IF LEN(sModemID) = 0 THEN
					// Same fallback the reference shell script uses. It is a
					// guess, and the router will reject it with 422 if wrong -
					// which at least says so clearly in sErrorText.
					sModemID := '1-1';
				END_IF
				uiStep := 30;
			END_IF

		ELSIF TON_Wait.Q THEN
			// Lookup timed out. Carry on with the fallback rather than failing
			// the whole job: the send step will report clearly if it is wrong.
			TON_Wait(IN := FALSE);
			fbCurl.curl_easy_abort();
			fbCurl.curl_slist_free_all(1);
			fbCurl.curl_easy_cleanup();
			sModemID := '1-1';
			uiStep   := 30;
		END_IF

	// -----------------------------------------------------------------
	30:	// SEND - start the request that actually delivers the message.
	// -----------------------------------------------------------------
		sStatus   := 'Steg 30: sender SMS...';
		sResponse := '';

		fbCurl.curl_easy_init();
		fbCurl.curl_set_RAM(ADR(sResponse), SIZEOF(sResponse));
		fbCurl.curl_easy_setopt_BOOL(64, FALSE);
		fbCurl.curl_easy_setopt_BOOL(81, FALSE);
		fbCurl.curl_easy_setopt_DINT(13, TIME_TO_DINT(tRequestTimeout) / 1000);
		fbCurl.curl_easy_setopt_DINT(78, 10);
		fbCurl.curl_easy_setopt_DINT(47, 1);

		sURL := CONCAT('https://', sRouterIP);
		sURL := CONCAT(sURL, '/api/messages/actions/send');
		fbCurl.curl_easy_setopt_STRING(10002, sURL);

		sHeader := CONCAT('Authorization: Bearer ', sToken);
		fbCurl.curl_slist_append(1, sHeader);
		fbCurl.curl_slist_append(1, 'Content-Type: application/json');
		fbCurl.curl_slist_append(1, 'Accept: */*');
		fbCurl.curl_easy_setopt_slist(10023, 1);
		// Some firmware versions refuse requests that carry no user agent.
		fbCurl.curl_easy_setopt_STRING(10018, 'curl/8.14.1');

		sBody := CONCAT('{"data":{"number":"', sNumber);
		sBody := CONCAT(sBody, '","message":"');
		sBody := CONCAT(sBody, sMessage);
		sBody := CONCAT(sBody, '","modem":"');
		sBody := CONCAT(sBody, sModemID);
		sBody := CONCAT(sBody, '"}}');
		fbCurl.curl_easy_setopt_STRING(10015, sBody);

		fbCurl.curl_easy_perform();
		TON_Wait(IN := FALSE);
		uiStep := 31;

	// -----------------------------------------------------------------
	31:	// SEND - wait for the router to accept or reject the message.
	//     This is the step where the duplicate question matters, because from
	//     here on the router may already have the message.
	// -----------------------------------------------------------------
		TON_Wait(IN := TRUE, PT := tWaitTimeout);
		IF fbCurl.xDone OR fbCurl.xError THEN
			TON_Wait(IN := FALSE);

			diHttpCode    := LINT_TO_DINT(fbCurl.curl_easy_getResponseCode());
			xCurlError    := fbCurl.xError;
			sCurlError    := fbCurl.sErrorString;
			sCurlSource   := fbCurl.sErrorSource;
			sLastResponse := LEFT(sResponse, 200);

			fbCurl.curl_slist_free_all(1);
			fbCurl.curl_easy_cleanup();

			IF FIND(sResponse, '"success":true') > 0 THEN
				uiStep := 100;

			ELSIF (diHttpCode = 401) AND NOT xRetriedLogin THEN
				// Refused token. A 401 proves the router did NOT take the
				// message, so logging in again and repeating cannot duplicate it.
				xTokenValid   := FALSE;
				sToken        := '';
				xRetriedLogin := TRUE;
				sStatus       := 'Token avvist - logger inn paa nytt';
				uiStep        := 10;

			ELSE
				// Drop the cached modem id so the next attempt looks it up
				// again. If the id was the problem, repeating it is pointless.
				sModemID   := '';
				sErrorText := CONCAT('Sending feilet, HTTP ', DINT_TO_STRING(diHttpCode));
				IF diHttpCode = 0 THEN
					// The request went out but nothing came back. The router may
					// already have queued the SMS, so the outcome is genuinely
					// unknown and the caller must not repeat it.
					xSendUncertain := TRUE;
					sErrorText := CONCAT(sErrorText, ' USIKKER curl: ');
					sErrorText := CONCAT(sErrorText, LEFT(sCurlError, 100));
				ELSE
					// A real HTTP answer reporting failure. Nothing was sent,
					// so the caller is free to try again.
					sErrorText := CONCAT(sErrorText, ' svar: ');
					sErrorText := CONCAT(sErrorText, LEFT(sResponse, 110));
				END_IF
				uiStep := 900;
			END_IF

		ELSIF TON_Wait.Q THEN
			// Aborted mid transfer. Same reasoning as above: the router may or
			// may not have taken it, so the message is flagged as uncertain.
			TON_Wait(IN := FALSE);
			fbCurl.curl_easy_abort();
			fbCurl.curl_slist_free_all(1);
			fbCurl.curl_easy_cleanup();
			xSendUncertain := TRUE;
			sModemID       := '';
			sErrorText     := 'Tidsavbrudd under sending - USIKKER, ikke send paa nytt';
			uiStep         := 900;
		END_IF

	// -----------------------------------------------------------------
	100: // DONE - the router confirmed the message.
	// -----------------------------------------------------------------
		xDone      := TRUE;
		xBusy      := FALSE;
		udiSentCnt := udiSentCnt + 1;
		tLastSend  := WagoAppTime.FuGetLocalDateAndTime();
		sStatus    := 'SMS sendt OK';
		uiStep     := 0;

	// -----------------------------------------------------------------
	900: // ERROR - sErrorText was filled in by whichever step failed.
	// -----------------------------------------------------------------
		xError      := TRUE;
		xBusy       := FALSE;
		udiErrorCnt := udiErrorCnt + 1;
		sStatus     := sErrorText;
		uiStep      := 0;

ELSE
	// Unknown step. Reached only if an online change moves the code under a
	// running state machine. Returning to idle is always safe.
	uiStep := 0;
END_CASE

(*
	ExtractJson                       Created 20.08.2026, rewritten 22.08.2026
	==========================================================================
	WHAT IT DOES
	Pulls the string value that belongs to a JSON key out of a raw HTTP answer.
	Used twice in this block: to lift the bearer token out of the login answer,
	and the modem id out of the modem status answer.

	HOW TO CALL IT
	sKey is the bare quoted key WITHOUT the colon, so the four characters that
	spell out id surrounded by quotes. The scanner then skips whatever separator
	follows, which means both of these parse correctly:
	    "id":"3-1"          compact
	    "id": "3-1"         with whitespace
	An empty string comes back when the key is not present, so the caller can
	simply test the length.

	*** WHY THIS IS A BYTE SCANNER AND NOT FIND AND MID ***
	The CODESYS standard string functions FIND, MID, LEFT and CONCAT are all
	declared with STRING(255) parameters. Handed a longer buffer they quietly
	look at the first 255 characters only, with no warning and no error.
	sResponse is STRING(4095). The login answer is short, so the token was
	always found and everything looked fine. But the modem status answer
	carries many fields per modem, and the id can sit past character 255 - so
	the lookup silently returned nothing, the block fell back to modem 1-1, and
	the router replied HTTP 422 Provided modem does not exist. Meanwhile the
	awk based shell script, which has no such limit, found 3-1 without trouble.

	This version walks the raw bytes through pointers instead, so the whole
	buffer is searched. The same approach is worth reaching for anywhere a long
	HTTP answer has to be parsed in ST.

	Character code 34 is the double quote, written numerically to keep the
	string literals in this method readable.
*)
METHOD ExtractJson : STRING(200)
VAR_INPUT
	sSource	: STRING(4095);		// Raw JSON body straight from the router
	sKey	: STRING(40);		// Quoted key to look for, without the colon
END_VAR
VAR
	pSrc	: POINTER TO BYTE;	// Walks sSource byte by byte
	pKey	: POINTER TO BYTE;	// Walks sKey during the comparison
	pRes	: POINTER TO BYTE;	// Writes into the result buffer
	iSrcLen	: INT;				// Real length of sSource, found by scanning for the terminator
	iKeyLen	: INT;				// Real length of sKey
	iPos	: INT;				// Current scan position in sSource
	iSub	: INT;				// Position inside the key while comparing
	iHit	: INT;				// Index just past the matched key. -1 means not found.
	iOut	: INT;				// Characters written to the result so far
	xMatch	: BOOL;				// Does the key match at the current position
	sResult	: STRING(200);		// Value being assembled, copied to the return at the end
END_VAR
// Default to empty, so every early exit below already returns the right thing.
ExtractJson := '';
sResult     := '';

pSrc := ADR(sSource);
pKey := ADR(sKey);
pRes := ADR(sResult);

// ---------------------------------------------------------------------
// Find the real lengths by scanning for the terminating zero. LEN cannot be
// used here for the same reason FIND cannot: it would stop at 255.
// Both loops are bounded by the declared buffer sizes, so a string that is
// somehow not terminated can never run off the end of memory.
// ---------------------------------------------------------------------
iKeyLen := 0;
WHILE (iKeyLen < 40) AND (pKey[iKeyLen] <> 0) DO
	iKeyLen := iKeyLen + 1;
END_WHILE
IF iKeyLen = 0 THEN
	RETURN;							// Nothing to search for
END_IF

iSrcLen := 0;
WHILE (iSrcLen < 4095) AND (pSrc[iSrcLen] <> 0) DO
	iSrcLen := iSrcLen + 1;
END_WHILE
IF iSrcLen < iKeyLen THEN
	RETURN;							// Answer is shorter than the key, so it cannot contain it
END_IF

// ---------------------------------------------------------------------
// Plain substring search across the whole buffer. Naive on purpose: the
// answers are a few kilobytes at most and this runs twice per message, so
// clarity is worth more here than a cleverer algorithm.
// ---------------------------------------------------------------------
iHit := -1;
iPos := 0;
WHILE (iPos <= (iSrcLen - iKeyLen)) AND (iHit < 0) DO
	xMatch := TRUE;
	iSub   := 0;
	WHILE (iSub < iKeyLen) AND xMatch DO
		IF pSrc[iPos + iSub] <> pKey[iSub] THEN
			xMatch := FALSE;		// Mismatch, stop comparing and slide along
		END_IF
		iSub := iSub + 1;
	END_WHILE
	IF xMatch THEN
		iHit := iPos + iKeyLen;		// First character after the key
	END_IF
	iPos := iPos + 1;
END_WHILE

IF iHit < 0 THEN
	RETURN;							// Key is not in this answer
END_IF

// ---------------------------------------------------------------------
// The next double quote after the key opens the value. Skipping forward to
// it rather than expecting a specific separator is what makes the parser
// tolerant of whitespace between the colon and the value.
// ---------------------------------------------------------------------
WHILE (iHit < iSrcLen) AND (pSrc[iHit] <> 34) DO
	iHit := iHit + 1;
END_WHILE
IF iHit >= iSrcLen THEN
	RETURN;							// No opening quote, so this is not a string value
END_IF
iHit := iHit + 1;					// Step onto the first character of the value itself

// ---------------------------------------------------------------------
// Copy until the closing quote. The output is capped at the size of the
// result buffer, and the terminator is written afterwards so the value is a
// valid IEC string whatever happens.
// ---------------------------------------------------------------------
iOut := 0;
WHILE (iHit < iSrcLen) AND (pSrc[iHit] <> 34) AND (iOut < 200) DO
	pRes[iOut] := pSrc[iHit];
	iOut       := iOut + 1;
	iHit       := iHit + 1;
END_WHILE
pRes[iOut] := 0;

ExtractJson := sResult;
END_METHOD

END_FUNCTION_BLOCK

// Teltonika/FbAlarmSlot
(*
	FbAlarmSlot                         Created 22.08.2026, rev 23.08.2026
	==========================================================================
	WHAT THIS BLOCK IS
	One alarm slot. It holds both the configuration for a single alarm and the
	live state of that alarm, and it does its own debouncing and edge detection.
	prg_AlarmSMS keeps an array of twenty of these.

	WHY A FUNCTION BLOCK AND NOT PARALLEL ARRAYS
	The CODESYS Best Practices for visualization recommend passing ONE parameter
	to a reusable visualization, ideally a function block instance, through
	VAR_IN_OUT so the instance is not copied. With one instance per alarm, a
	frame that shows one row needs a single reference:

	    alarm  ->  prg_AlarmSMS.aAlarm[7]

	instead of one reference per field. The same document also advises keeping
	object state inside the function block rather than in the visualization,
	which is why the debounce timer and the edge memory live here.

	EVERYTHING THE OPERATOR EDITS IS AN INPUT
	A visualization can only write to VAR_INPUT and VAR_IN_OUT. Outputs are
	display only. That is the reason the delay is entered as iDelaySec rather
	than as the TIME value itself, and the reason the recipient selection is a
	plain array of BOOL rather than a bit mask: a checkbox binds straight to
	axToRecipient[2] with no bit arithmetic anywhere.

	HOW IT IS USED
	Call the instance once per cycle with no arguments:

	    aAlarm[i]();
	    IF aAlarm[i].xRising THEN ... send an alarm message ... END_IF
*)
FUNCTION_BLOCK FbAlarmSlot
VAR_INPUT
	// === CONFIGURATION - written by the operator, usually from a visualization ===

	xSmsEnable	: BOOL  := FALSE;		// The on and off switch for this alarm. TRUE means it is
										// allowed to send an SMS, FALSE means it is still tracked
										// but stays silent. Bind a CHECKBOX to this, not a radio
										// button: each alarm is independent of the others.

	sText		: STRING(70) := '';		// The wording that ends up in the message. Keep it short:
										// the site name and time stamp are added in front, and the
										// total is capped at 140 characters. Avoid double quotes -
										// the sender replaces them with spaces so they cannot break
										// the JSON body.

	// Which of the four phone numbers this alarm goes to. One BOOL per person,
	// so a visualization binds four independent CHECKBOX elements:
	//     alarm.axToRecipient[1]   ... alarm.axToRecipient[4]
	// Radio buttons are wrong here - they are mutually exclusive, and one alarm
	// must be able to reach several people at once.
	// The size is fixed at four and must match MAX_RECIPIENTS in the program.
	axToRecipient : ARRAY[1..4] OF BOOL := [TRUE, FALSE, FALSE, FALSE];

	iDelaySec	: INT   := 30;			// Debounce time in SECONDS. How long xAlarmIn must stay
										// TRUE before it counts as a real alarm, which filters out
										// flicker and short network dropouts. This is the single
										// biggest contributor to the delay between a fault
										// appearing and the SMS arriving.
										// Seconds rather than minutes because some alarms need to
										// react inside a minute: 30 is thirty seconds, 300 is five
										// minutes. The block clamps the value to a sane range and
										// shows it back in readable form through sDelayText.

	// === PLANT SIGNAL - written by whatever logic detects the condition ===

	xAlarmIn	: BOOL;					// The raw alarm condition, TRUE means the fault is present.
										// Write it from anywhere in the project, for example:
										//   prg_AlarmSMS.aAlarm[1].xAlarmIn := NOT xPriceDataValid;
END_VAR
VAR_OUTPUT
	// === LIVE STATE - read only, produced by this block ===

	xActive		: BOOL;					// The debounced alarm state. This is the one to show on a
										// lamp, because it matches what the SMS logic reacts to.
										// xAlarmIn may flicker; xActive does not.

	xRising		: BOOL;					// TRUE for exactly one call, on the cycle where the alarm
										// became active. The owner uses this to send one message
										// rather than one per cycle for as long as the fault lasts.

	xFalling	: BOOL;					// TRUE for exactly one call, on the cycle where the alarm
										// cleared. Used for the optional message that tells the
										// operator the fault went away.

	tOnDelay	: TIME;					// iDelaySec expressed as a TIME, which is what the timer
										// actually uses. Read only: change the delay through
										// iDelaySec, not here.

	sDelayText	: STRING(12);			// The delay rendered for a screen, for example 30 s or
										// 5 min. Bind a text field to this with the %s placeholder.
END_VAR
VAR
	TON_Delay	: TON;					// Implements the debounce. Held here rather than in the
										// caller so every alarm carries its own timing with it.
	xPrev		: BOOL;					// Previous value of xActive, so the two edge outputs can be
										// derived. Without it a standing alarm would keep firing.
END_VAR
VAR CONSTANT
	DELAY_MAX_SEC : INT := 3600;		// One hour. An upper bound so a mistyped value in the
										// visualization cannot mute an alarm for days.
END_VAR

// =====================================================================
// Turn the operator setting into the value the timer needs.
// The visualization writes whole seconds into iDelaySec, because a text
// field cannot write a TIME and the %d placeholder on a TIME would show raw
// milliseconds. Clamping happens here so a typing mistake in the screen can
// never produce a negative time or mute an alarm for days.
// =====================================================================
IF iDelaySec < 0 THEN
	iDelaySec := 0;
ELSIF iDelaySec > DELAY_MAX_SEC THEN
	iDelaySec := DELAY_MAX_SEC;
END_IF

tOnDelay := UDINT_TO_TIME(INT_TO_UDINT(iDelaySec) * 1000);

// Readable version for the screen. Whole minutes above a minute, seconds
// below it. Any remaining seconds are dropped on purpose: the field is a
// quick overview, and the exact value is always visible in iDelaySec.
IF iDelaySec < 60 THEN
	sDelayText := CONCAT(INT_TO_STRING(iDelaySec), ' s');
ELSE
	sDelayText := CONCAT(INT_TO_STRING(iDelaySec / 60), ' min');
END_IF

// =====================================================================
// Debounce.
// The timer only reaches Q once the raw signal has been TRUE continuously
// for tOnDelay. A signal that drops out in the meantime restarts it, so a
// brief glitch never becomes a text message in the middle of the night.
// =====================================================================
TON_Delay(IN := xAlarmIn, PT := tOnDelay);
xActive := TON_Delay.Q;

// =====================================================================
// Edge detection on the DEBOUNCED state, not on the raw input.
// Both outputs are true for a single call only. Deriving them here means the
// caller never has to keep its own edge memory, and cannot get it wrong.
// =====================================================================
xRising  := xActive AND NOT xPrev;
xFalling := (NOT xActive) AND xPrev;

// Remember the state for the next call. This runs unconditionally: even when
// the alarm is muted its state must keep tracking, otherwise unmuting it
// later would produce a false edge for a fault that was already standing.
xPrev := xActive;

END_FUNCTION_BLOCK

// /AlarmAlarms
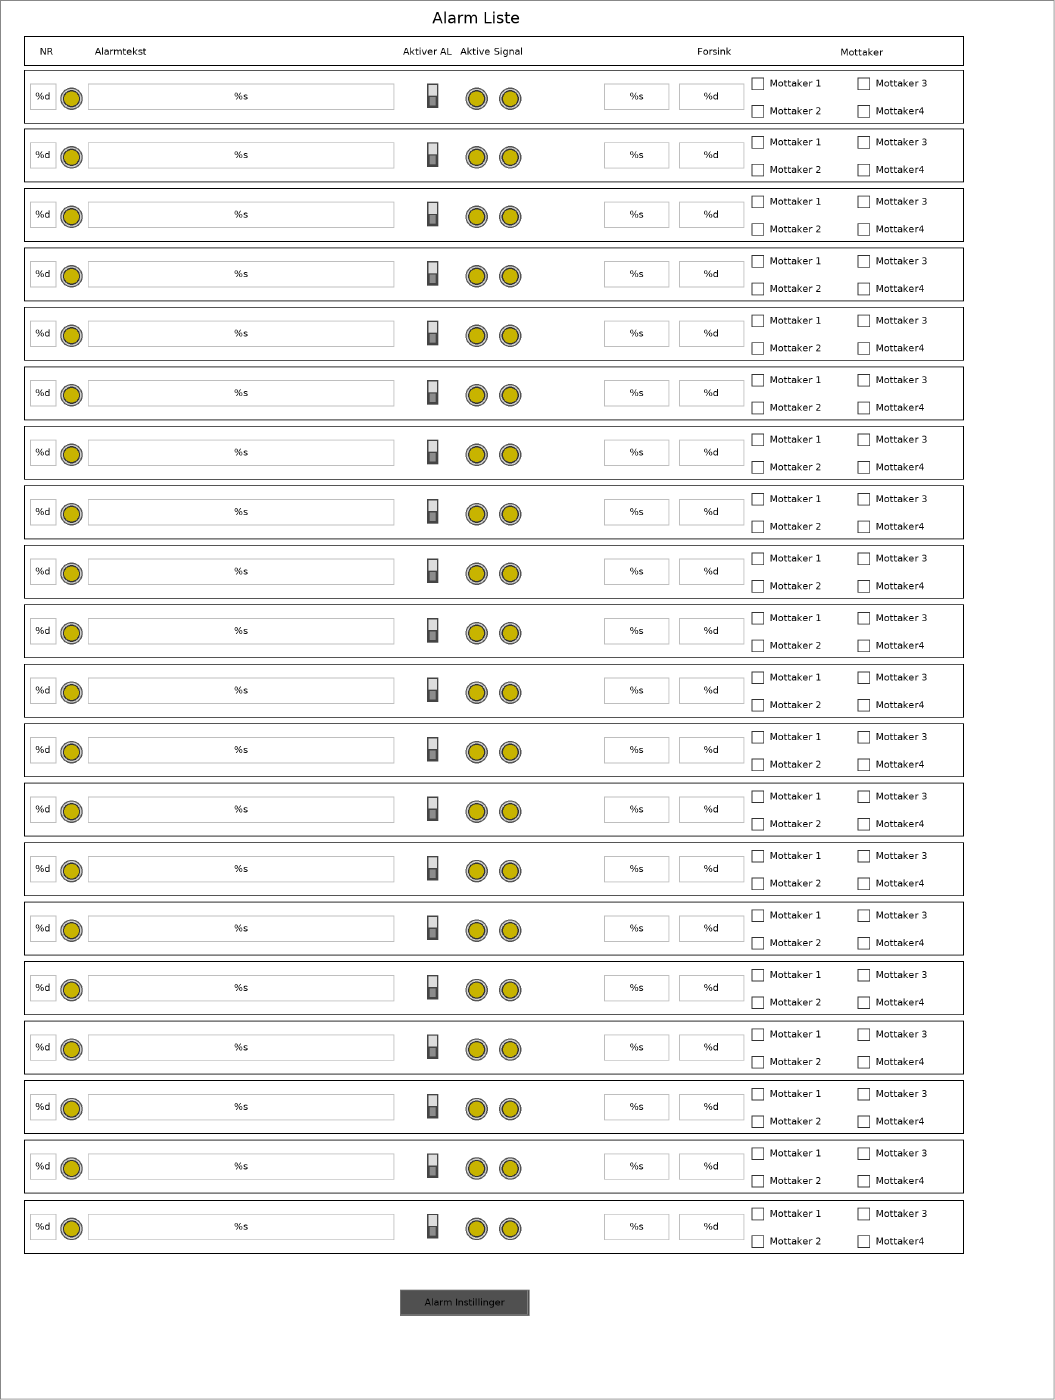
VISUALIZATION AlarmAlarms  // 1224x1624
    RoundedRectangle (28,42 1090x34)
    Label (34,45 40x30), "NR"
    Label (102,45 76x30), "Alarmtekst"
    Label (459,45 70x30), "Aktiver AL"
    Label (528,45 47x30), "Aktive"
    Label (965,46 70x30), "Mottaker"
    Label (794,45 70x30), "Forsink"
    Frame (28,81 1090x62)
        shows AlarmerListe(alarm := prg_AlarmSMS.aAlarm[1], iNr := 1)
    Frame (28,149 1090x62)
        shows AlarmerListe(alarm := prg_AlarmSMS.aAlarm[2], iNr := 2)
    Frame (28,218 1090x62)
        shows AlarmerListe(alarm := prg_AlarmSMS.aAlarm[3], iNr := 3)
    Frame (28,287 1090x62)
        shows AlarmerListe(alarm := prg_AlarmSMS.aAlarm[4], iNr := 4)
    Frame (28,356 1090x62)
        shows AlarmerListe(alarm := prg_AlarmSMS.aAlarm[5], iNr := 5)
    Frame (28,425 1090x62)
        shows AlarmerListe(alarm := prg_AlarmSMS.aAlarm[6], iNr := 6)
    Frame (28,494 1090x62)
        shows AlarmerListe(alarm := prg_AlarmSMS.aAlarm[7], iNr := 7)
    Frame (28,563 1090x62)
        shows AlarmerListe(alarm := prg_AlarmSMS.aAlarm[8], iNr := 8)
    Frame (28,632 1090x62)
        shows AlarmerListe(alarm := prg_AlarmSMS.aAlarm[9], iNr := 9)
    Frame (28,701 1090x62)
        shows AlarmerListe(alarm := prg_AlarmSMS.aAlarm[10], iNr := 10)
    Frame (28,770 1090x62)
        shows AlarmerListe(alarm := prg_AlarmSMS.aAlarm[11], iNr := 11)
    Frame (28,839 1090x62)
        shows AlarmerListe(alarm := prg_AlarmSMS.aAlarm[12], iNr := 12)
    Frame (28,908 1090x62)
        shows AlarmerListe(alarm := prg_AlarmSMS.aAlarm[13], iNr := 13)
    Frame (28,977 1090x62)
        shows AlarmerListe(alarm := prg_AlarmSMS.aAlarm[14], iNr := 14)
    Frame (28,1046 1090x62)
        shows AlarmerListe(alarm := prg_AlarmSMS.aAlarm[15], iNr := 15)
    Frame (28,1115 1090x62)
        shows AlarmerListe(alarm := prg_AlarmSMS.aAlarm[16], iNr := 16)
    Frame (28,1184 1090x62)
        shows AlarmerListe(alarm := prg_AlarmSMS.aAlarm[17], iNr := 17)
    Frame (28,1253 1090x62)
        shows AlarmerListe(alarm := prg_AlarmSMS.aAlarm[18], iNr := 18)
    Frame (28,1322 1090x62)
        shows AlarmerListe(alarm := prg_AlarmSMS.aAlarm[19], iNr := 19)
    Frame (28,1392 1090x62)
        shows AlarmerListe(alarm := prg_AlarmSMS.aAlarm[20], iNr := 20)
    Label (566,45 48x30), "Signal"
    Label (454,6 197x30), "Alarm Liste"
    Button (464,1496 150x30), "Alarm Instillinger"
        OnMouseClick:  Assign=AlarmMain, Type=Assignment
END_VISUALIZATION

// /AlarmerListe
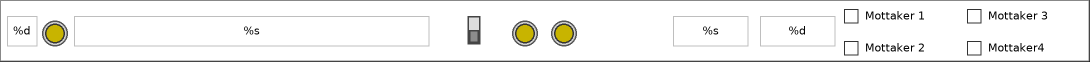
VISUALIZATION AlarmerListe  // 1090x62
VAR_IN_OUT
    alarm : FbAlarmSlot;
END_VAR
VAR_INPUT
    iNr : INT;
END_VAR
    RoundedRectangle (0,0 1090x62)
    Textfield (7,16 30x30), "%d", text variable: iNr
    Textfield (74,16 355x30), "%s", text variable: alarm.sText
        OnMouseClick: write alarm.sText via Edit
    Lamp1 (510,16 30x35), variable: alarm.xActive, style: Lamp-Lamp1-Yellow
    Textfield (673,16 75x30), "%s", text variable: alarm.sDelayText
    Lamp1 (549,16 30x35), variable: alarm.xAlarmIn, style: Lamp-Lamp1-Yellow
    Textfield (760,16 75x30), "%d", text variable: alarm.iDelaySec
        OnMouseClick: write alarm.iDelaySec via Default, min 0, max 3600
    DipSwitch (439,16 70x28), variable: alarm.xSmsEnable, behaviour: TOGGLE, style: Switch-DipSwitch-Gray
    Lamp1 (40,16 30x35), variable: alarm.xSmsEnable, style: Lamp-Lamp1-Yellow
    Checkbox (842,1 107x30), "Mottaker 1", variable: alarm.axToRecipient[1]
    Checkbox (842,33 107x30), "Mottaker 2", variable: alarm.axToRecipient[2]
    Checkbox (965,33 107x30), "Mottaker4", variable: alarm.axToRecipient[4]
    Checkbox (965,1 107x30), "Mottaker 3", variable: alarm.axToRecipient[3]
END_VISUALIZATION

// /AlarmMain
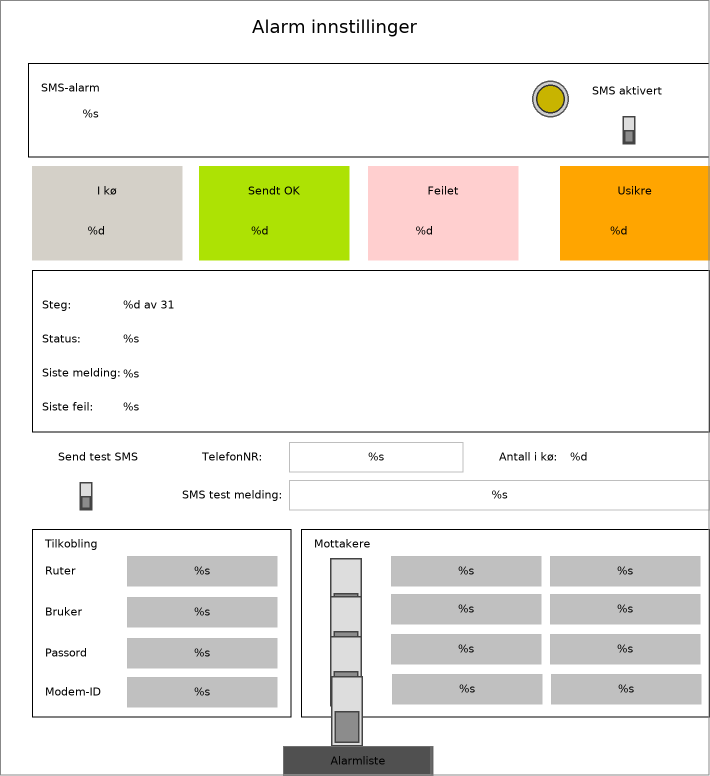
VISUALIZATION AlarmMain  // 710x776
    RoundedRectangle (28,63 681x94)
    Label (38,73 77x30), "SMS-alarm"
    Textfield (42,99 97x30), "%s", text variable: prg_AlarmSMS.sSiteName
    Lamp1 (529,76 43x46), variable: prg_AlarmSMS.xSmsGlobalEnable, style: Lamp-Lamp1-Yellow
    Label (582,76 90x30), "SMS aktivert"
    RoundedRectangle (32,166 150x94)
    Label (32,176 150x30), "I kø"
    Textfield (39,216 115x30), "%d", text variable: prg_AlarmSMS.iQueueCount
    DipSwitch (594,116 70x28), variable: prg_AlarmSMS.xSmsGlobalEnable, behaviour: TOGGLE, style: Switch-DipSwitch-Gray
    RoundedRectangle (199,166 150x94)
    Label (199,176 150x30), "Sendt OK"
    Textfield (206,216 108x30), "%d", text variable: prg_AlarmSMS.udiSentOk
    RoundedRectangle (368,166 150x94)
    Label (368,176 150x30), "Feilet"
    Textfield (368,216 113x30), "%d", text variable: prg_AlarmSMS.udiSendFailed
    RoundedRectangle (560,166 150x94)
    Label (560,176 150x30), "Usikre"
    Textfield (567,216 104x30), "%d", text variable: prg_AlarmSMS.udiUncertain
    RoundedRectangle (32,270 678x162)
    Label (39,290 90x30), "Steg:"
    Textfield (120,290 560x30), "%d av 31", text variable: prg_AlarmSMS.uiSendStep
    Textfield (120,324 560x30), "%s", text variable: prg_AlarmSMS.sSmsStatus
    Label (39,324 90x30), "Status:"
    Label (39,358 90x30), "Siste melding:"
    Textfield (120,359 560x30), "%s", text variable: prg_AlarmSMS.sLastMessage
    Textfield (120,392 560x30), "%s", text variable: prg_AlarmSMS.sLastError
    Label (39,392 90x30), "Siste feil:"
    Label (39,442 118x30), "Send test SMS"
    DipSwitch (51,482 70x28), variable: prg_AlarmSMS.xManualSend, behaviour: TOGGLE, style: Switch-DipSwitch-Gray
    Label (173,442 118x30), "TelefonNR:"
    Label (173,480 118x30), "SMS test melding:"
    Textfield (289,442 174x30), "%s", text variable: prg_AlarmSMS.sTestNumber
        OnMouseClick: write the text variable via Edit
    Textfield (289,480 421x30), "%s", text variable: prg_AlarmSMS.sManualText
        OnMouseClick: write the text variable via Edit
    RoundedRectangle (32,529 259x188)
    Label (42,529 73x30), "Tilkobling"
    Label (42,556 44x30), "Ruter"
    Label (42,597 58x30), "Bruker"
    Label (42,638 84x30), "Passord"
    Label (42,677 84x30), "Modem-ID"
    Textfield (127,556 150x30), "%s", text variable: prg_AlarmSMS.sRouterOverride
        OnMouseClick: write the text variable via Edit
    Textfield (127,597 150x30), "%s", text variable: GVL_TeltonikaCredentials.Teltonika_Username
        OnMouseClick: write the text variable via Edit
    Textfield (127,638 150x30), "%s", text variable: GVL_TeltonikaCredentials.Teltonika_Password
        OnMouseClick: write the text variable via Edit
    Textfield (127,677 150x30), "%s", text variable: prg_AlarmSMS.sModemIdForced
        OnMouseClick: write the text variable via Edit
    RoundedRectangle (301,529 409x188)
    Label (311,529 73x30), "Mottakere"
    DipSwitch (311,558 70x70), variable: prg_AlarmSMS.axRecipientEnable[1], behaviour: TOGGLE, style: Switch-DipSwitch-Gray
    Textfield (391,556 150x30), "%s", text variable: prg_AlarmSMS.asRecipientName[1]
        OnMouseClick: write the text variable via Edit
    Textfield (550,556 150x30), "%s", text variable: prg_AlarmSMS.asRecipientNumber[1]
        OnMouseClick: write the text variable via Edit
    DipSwitch (311,596 70x70), variable: prg_AlarmSMS.axRecipientEnable[2], behaviour: TOGGLE, style: Switch-DipSwitch-Gray
    Textfield (391,594 150x30), "%s", text variable: prg_AlarmSMS.asRecipientName[2]
        OnMouseClick: write the text variable via Edit
    Textfield (550,594 150x30), "%s", text variable: prg_AlarmSMS.asRecipientNumber[2]
        OnMouseClick: write the text variable via Edit
    DipSwitch (311,636 70x70), variable: prg_AlarmSMS.axRecipientEnable[3], behaviour: TOGGLE, style: Switch-DipSwitch-Gray
    Textfield (391,634 150x30), "%s", text variable: prg_AlarmSMS.asRecipientName[3]
        OnMouseClick: write the text variable via Edit
    Textfield (550,634 150x30), "%s", text variable: prg_AlarmSMS.asRecipientNumber[3]
        OnMouseClick: write the text variable via Edit
    DipSwitch (312,676 70x70), variable: prg_AlarmSMS.axRecipientEnable[4], behaviour: TOGGLE, style: Switch-DipSwitch-Gray
    Textfield (392,674 150x30), "%s", text variable: prg_AlarmSMS.asRecipientName[4]
        OnMouseClick: write the text variable via Edit
    Textfield (551,674 150x30), "%s", text variable: prg_AlarmSMS.asRecipientNumber[4]
        OnMouseClick: write the text variable via Edit
    Label (496,442 67x30), "Antall i kø:"
    Textfield (560,442 38x30), "%d", text variable: prg_AlarmSMS.iTestQueued
    Button (283,746 150x30), "Alarmliste"
        OnMouseClick:  Assign=AlarmAlarms, Type=Assignment
    Label (236,12 197x30), "Alarm innstillinger"
END_VISUALIZATION
